Fanuc KAREL source: IO0012.KL

PROGRAM IO0012
%NOLOCKGROUP
ROUTINE RTEST
VAR
  I : INTEGER
  STATUS : INTEGER
  ENTRY : INTEGER
  A : ARRAY[3] OF INTEGER
  B : BOOLEAN
  R : REAL
  P : XYZWPR
  JPOS : JOINTPOS
  PF : POSITION
BEGIN
  I = 1
  A[1] = 2
  B = TRUE
  R = 1.0
  WAIT FOR DIN[I + 1] = ON
END RTEST
BEGIN
  RTEST
END IO0012
